TYPE E_JobType :
(
	E_JobType_MoveStone,
	E_JobType_NewStone,
	E_JobType_RemoveStone
);
END_TYPE

(* stored: Version 1.1.0.1, ProductVersion 3.1.4024.9
   DUT E_JobType: Id {3a28bf40-c80a-4ed1-9bcd-c95db6d216cd} *)
